FUNCTION_BLOCK FB_MotorBase IMPLEMENTS I_Motor
VAR_OUTPUT
    updates : UDINT;
    bodyCalls : UDINT;
END_VAR
VAR
    speed : LREAL := 0.5;
    runningState : BOOL;
END_VAR

bodyCalls := bodyCalls + 1;

METHOD PUBLIC Update
VAR_INPUT
    run : BOOL;
    delay : TIME;
END_VAR
VAR_INST
    startup : TON;
END_VAR
updates := updates + 1;
(* The protected property reaches the most-derived CheckFault hook. *)
startup(IN := run AND THIS^.MayRun, PT := delay);
THIS^.runningState := startup.Q;
END_METHOD

METHOD PROTECTED CheckFault : BOOL
CheckFault := FALSE;
END_METHOD

METHOD PRIVATE ClampSpeed : LREAL
VAR_INPUT
    value : LREAL;
END_VAR
ClampSpeed := LIMIT(0.0, value, 1.0);
END_METHOD

PROPERTY PROTECTED MayRun : BOOL
GET
MayRun := NOT THIS^.CheckFault();
END_GET
END_PROPERTY

PROPERTY PUBLIC SpeedSetpoint : LREAL
GET
SpeedSetpoint := THIS^.speed;
END_GET
SET
THIS^.speed := THIS^.ClampSpeed(value := SpeedSetpoint);
END_SET
END_PROPERTY

PROPERTY PUBLIC Running : BOOL
GET
Running := THIS^.runningState;
END_GET
END_PROPERTY

PROPERTY PUBLIC Faulted : BOOL
GET
Faulted := THIS^.CheckFault();
END_GET
END_PROPERTY

PROPERTY PUBLIC ActualSpeed : LREAL
GET
IF THIS^.runningState THEN
    ActualSpeed := THIS^.speed;
ELSE
    ActualSpeed := 0.0;
END_IF;
END_GET
END_PROPERTY

END_FUNCTION_BLOCK

(* stored: Version 1.1.0.1, ProductVersion 3.1 *)
